Fanuc KAREL source: kt00036.KL

-- PROVISIONAL review KL for V1013-1; original PC SHA256 8ce9b10fd524e722409ba41dbf9be3229b6ae66c1b20fc2665798d928c88af58
-- Incomplete behavior may be omitted. Consult companion uncertainty JSON. Do not deploy.
PROGRAM KT00036
%NOLOCKGROUP
VAR
  I1 : INTEGER
  R2 : REAL
  OUT : REAL
BEGIN
  -- UNRESOLVED_PC offsets 5-16; opcodes 2E,23
  -- UNRESOLVED_PC offsets 21-32; opcodes 2E,23
  -- UNRESOLVED_PC offsets 37-59; opcodes 21,21,29,64,29,6A,23
  -- UNRESOLVED_PC offsets 64-68; opcodes 7F
END KT00036
